FUNCTION_BLOCK Controle_Revezamento_3 (* Revezamento de 3 equipamentos por tempo como principal (padrao Revezamento_3_Motores do legado) *)
  (* Standard: 61499-2 *)
  (* Version 1.0, 21/10/2026, Hidryco, Hidryco, 1.0: Revezamento de 3 equipamentos por tempo como principal (padrao Revezamento_3_Motores do legado) *)
  PACKAGE Hidryco.HidrycoLib;
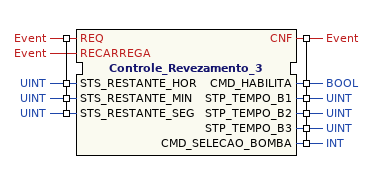
  EVENT_INPUT
    REQ WITH STS_RESTANTE_HOR, STS_RESTANTE_MIN, STS_RESTANTE_SEG; (* Status vindo do processo *)
    RECARREGA; (* Reenvia os ajustes persistentes (chamado no fim do INIT do processo) *)
  END_EVENT
  EVENT_OUTPUT
    CNF WITH CMD_HABILITA, STP_TEMPO_B1, STP_TEMPO_B2, STP_TEMPO_B3, CMD_SELECAO_BOMBA; (* Ajustes para o processo (mudanca na IHM, OPC UA ou recarga) *)
  END_EVENT
  VAR_INPUT
    STS_RESTANTE_HOR : UINT; (* Tempo para a troca da principal (h) *)
    STS_RESTANTE_MIN : UINT; (* Tempo para a troca da principal (min) *)
    STS_RESTANTE_SEG : UINT; (* Tempo para a troca da principal (s) *)
  END_VAR
  VAR_OUTPUT
    CMD_HABILITA : BOOL; (* Troca da principal por tempo *)
    STP_TEMPO_B1 : UINT; (* Horas do equipamento 1 como principal *)
    STP_TEMPO_B2 : UINT; (* Horas do equipamento 2 como principal *)
    STP_TEMPO_B3 : UINT; (* Horas do equipamento 3 como principal *)
    CMD_SELECAO_BOMBA : INT; (* Bomba principal *)
  END_VAR
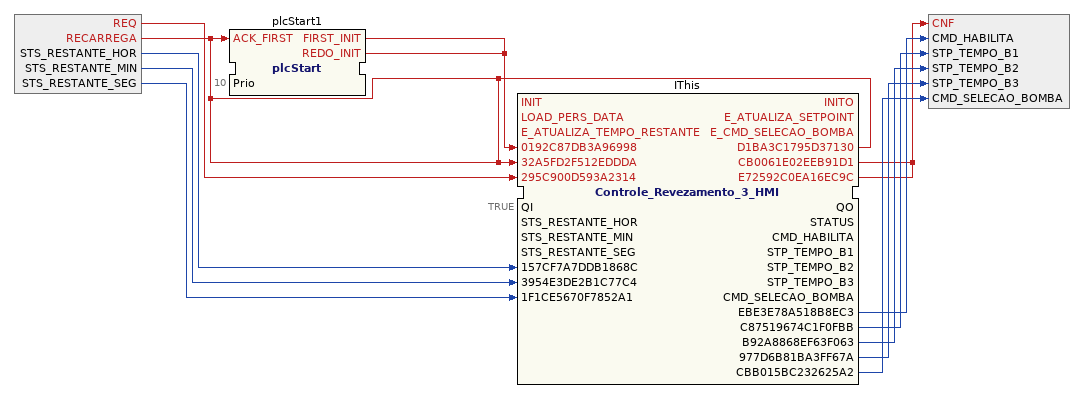
  FBS
    IThis : Controle_Revezamento_3_HMI(QI := TRUE);
    plcStart1 : plcStart(Prio := 10);
  END_FBS
  EVENT_CONNECTIONS
    plcStart1.FIRST_INIT TO IThis.0192C87DB3A96998;
    plcStart1.REDO_INIT TO IThis.0192C87DB3A96998;
    IThis.D1BA3C1795D37130 TO IThis.32A5FD2F512EDDDA;
    IThis.D1BA3C1795D37130 TO plcStart1.ACK_FIRST;
    RECARREGA TO IThis.32A5FD2F512EDDDA;
    IThis.CB0061E02EEB91D1 TO CNF;
    IThis.E72592C0EA16EC9C TO CNF;
    REQ TO IThis.295C900D593A2314;
  END_CONNECTIONS
  DATA_CONNECTIONS
    IThis.EBE3E78A518B8EC3 TO CMD_HABILITA;
    IThis.C87519674C1F0FBB TO STP_TEMPO_B1;
    IThis.B92A8868EF63F063 TO STP_TEMPO_B2;
    IThis.977D6B81BA3FF67A TO STP_TEMPO_B3;
    IThis.CBB015BC232625A2 TO CMD_SELECAO_BOMBA;
    STS_RESTANTE_HOR TO IThis.157CF7A7DDB1868C;
    STS_RESTANTE_MIN TO IThis.3954E3DE2B1C77C4;
    STS_RESTANTE_SEG TO IThis.1F1CE5670F7852A1;
  END_CONNECTIONS
END_FUNCTION_BLOCK
